FUNCTION_BLOCK F (* Negative C4: a CASE on arithmetic over the position, in an algorithm shared by two control states *)
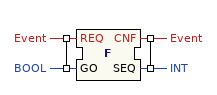
  EVENT_INPUT
    REQ WITH GO;
  END_EVENT
  EVENT_OUTPUT
    CNF WITH SEQ;
  END_EVENT
  VAR_INPUT
    GO : BOOL;
  END_VAR
  VAR_OUTPUT
    SEQ : INT;
  END_VAR
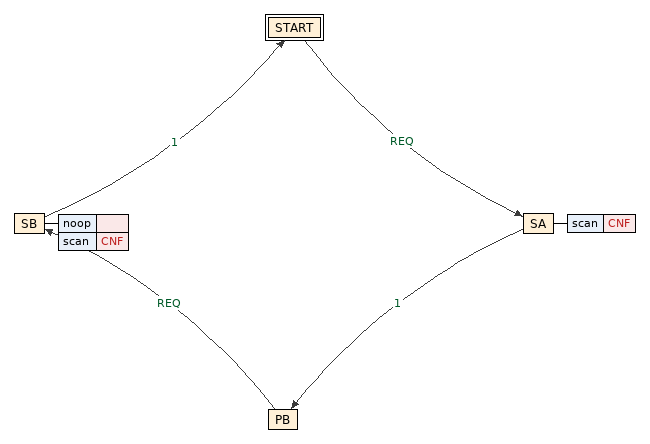
  EC_STATES
    START;
    SA : scan -> CNF;
    PB;
    SB : noop, scan -> CNF;
  END_STATES
  EC_TRANSITIONS
    START TO SA := REQ;
    SA TO PB := 1;
    PB TO SB := REQ;
    SB TO START := 1;
  END_TRANSITIONS
  ALGORITHM scan IN ST:
CASE SEQ + 0 OF
  0:
    IF GO THEN
      SEQ := 1;
    END_IF;
  1:
    SEQ := 2;
  2:
    SEQ := 0;
END_CASE;
  END_ALGORITHM
  ALGORITHM noop IN ST:
SEQ := SEQ;
  END_ALGORITHM
END_FUNCTION_BLOCK
